// FB_CTUD: 加减计数器
// 描述: CU上升沿加1, CD上升沿减1

FUNCTION_BLOCK FB_CTUD
VAR_INPUT
    CU  : BOOL;   // 加计数脉冲输入 (上升沿有效)
    CD  : BOOL;   // 减计数脉冲输入 (上升沿有效)
    R   : BOOL;   // 复位输入 (TRUE时CV=0)
    LOAD: BOOL;   // 加载输入 (TRUE时CV=PV)
    PV  : INT;    // 预设计数值
END_VAR
VAR_OUTPUT
    QU  : BOOL;   // 加计数完成输出 (CV>=PV)
    QD  : BOOL;   // 减计数完成输出 (CV<=0)
    CV  : INT;    // 当前计数值
END_VAR
VAR
    LastCU : BOOL := FALSE;
    LastCD : BOOL := FALSE;
END_VAR

BEGIN
    // R为TRUE时复位
    IF #R THEN
        #CV := 0;
    ELSIF #LOAD THEN
        // LOAD为TRUE时加载PV
        #CV := #PV;
    ELSE
        // CU上升沿且CV<PV时加1
        IF #CU AND NOT #LastCU THEN
            IF #CV < #PV THEN
                #CV := #CV + 1;
            END_IF;
        END_IF;

        // CD上升沿且CV>0时减1
        IF #CD AND NOT #LastCD THEN
            IF #CV > 0 THEN
                #CV := #CV - 1;
            END_IF;
        END_IF;
    END_IF;

    // 更新输出状态
    #QU := (#CV >= #PV);
    #QD := (#CV <= 0);

    #LastCU := #CU;
    #LastCD := #CD;

END_FUNCTION_BLOCK
